(* IEC 61131-3 sources: axsharp/src/tests.integrations/integrated/src/ax/src/dataswapping, 4 files *)

(* ---- myEnum.st ---- *)
TYPE myEnum :
    (
        Unknown,
        Available,
        UnAvailable
    );
    END_TYPE

(* ---- all_primitives.st ---- *)
{S7.extern=ReadWrite}
CLASS all_primitives
    VAR PUBLIC
        myBOOL	        :       BOOL	      ;
        myBYTE	        :       BYTE	      ;
        myWORD	        :       WORD	      ;
        myDWORD	        :       DWORD	      ;
        myLWORD	        :       LWORD	      ;
        mySINT	        :       SINT	      ;
        myINT	        :       INT	          ;
        myDINT	        :       DINT	      ;
        myLINT	        :       LINT	      ;
        myUSINT	        :       USINT	      ;
        myUINT	        :       UINT	      ;
        myUDINT	        :       UDINT	      ;
        myULINT	        :       ULINT	      ;
        myREAL	        :       REAL	      ;
        myLREAL	        :       LREAL	      ;
        myTIME	        :       TIME	      ;
        myLTIME	        :       LTIME	      ;
        myDATE	        :       DATE	      ;
     //   myLDATE	        :       LDATE	      ;
        myTIME_OF_DAY	:       TIME_OF_DAY	  ;
     //   myLTIME_OF_DAY	:       LTIME_OF_DAY  ;
        myDATE_AND_TIME  :      DATE_AND_TIME ;
     //   myLDATE_AND_TIME :      LDATE_AND_TIME;
     //   myCHAR	        :       CHAR	      ;
     //   myWCHAR	        :       WCHAR	      ;
        mySTRING	        :   STRING	      ;
        myWSTRING	    :       WSTRING	      ;
        myEnum : myEnum;
    END_VAR

END_CLASS

(* ---- moster.st ---- *)
NAMESPACE MonsterData
    {S7.extern=ReadWrite}
    CLASS MonsterBase
        VAR PUBLIC
            Description : STRING;
            Id : ULINT;
            ArrayOfBytes : ARRAY[0..3] OF BYTE;
            ArrayOfDrives : ARRAY[0..3] OF DriveBase;

            {#ix-attr:[IgnoreOnPocoOperation()]}
            DriveBase_tobeignoredbypocooperations : DriveBase;

            {#ix-attr:[IgnoreOnPocoOperation()]}
            Description_tobeignoredbypocooperations : STRING;
        END_VAR
    END_CLASS
    {S7.extern=ReadWrite}
    CLASS Monster EXTENDS MonsterBase
        VAR PUBLIC
            DriveA : DriveBase;
        END_VAR
    END_CLASS

    {S7.extern=ReadWrite}
    CLASS DriveBase
        VAR PUBLIC
            Position : LREAL;
            Velo : LREAL;
            Acc : LREAL;
            Dcc : LREAL;
        END_VAR
    END_CLASS
END_NAMESPACE

(* ---- realmonster.st ---- *)
NAMESPACE RealMonsterData
    {S7.extern=ReadWrite}
    CLASS RealMonsterBase
        VAR PUBLIC
            Description : STRING;
            Id : ULINT;
            TestDate : DATE;
            TestDateTime: DATE_AND_TIME;
            TestTimeSpan: TIME_OF_DAY;
            ArrayOfBytes : ARRAY[0..3] OF BYTE;
            ArrayOfDrives : ARRAY[0..3] OF DriveBaseNested;
        END_VAR
    END_CLASS

    {S7.extern=ReadWrite}
    CLASS RealMonster EXTENDS RealMonsterBase
        VAR PUBLIC
            DriveA : DriveBaseNested;
        END_VAR
    END_CLASS

    {S7.extern=ReadWrite}
    CLASS DriveBaseNested
        VAR PUBLIC
            Position : LREAL;
            Velo : LREAL;
            Acc : LREAL;
            Dcc : LREAL;
            NestedLevelOne : NestedLevelOne;
        END_VAR
    END_CLASS

    {S7.extern=ReadWrite}
    CLASS NestedLevelOne
        VAR PUBLIC
            Position : LREAL;
            Velo : LREAL;
            Acc : LREAL;
            Dcc : LREAL;
            NestedLevelTwo: NestedLevelTwo;
        END_VAR
    END_CLASS

    {S7.extern=ReadWrite}
    CLASS NestedLevelTwo
        VAR PUBLIC
            Position : LREAL;
            Velo : LREAL;
            Acc : LREAL;
            Dcc : LREAL;
            NestedLevelThree: NestedLevelThree;
        END_VAR
    END_CLASS

    {S7.extern=ReadWrite}
    CLASS NestedLevelThree
        VAR PUBLIC
            Position : LREAL;
            Velo : LREAL;
            Acc : LREAL;
            Dcc : LREAL;
        END_VAR
    END_CLASS

END_NAMESPACE
